Fanuc KAREL source: KO00035.KL

PROGRAM KO00035
%NOLOCKGROUP
%ENVIRONMENT MIR
VAR
  P1: POSITION
  P2: POSITION
  F: BOOLEAN
  OUT: XYZWPREXT
BEGIN
  F = TRUE
  OUT = MIRROR(P1, P2, F)
END KO00035
